(* IEC 61131-3 sources: iolistgen/src/POUs/PRG_Main, 2 files *)

(* ---- PRG_Main.decl.st ---- *)
// Назначение: точка входа приложения проверки сгенерированного кода (пример КНС-1, examples/kns): логика
//             станции в минимальном объёме — регулятор уровня LIC101 (тип Pid: вызов пишет логика станции,
//             контракт plc-process-lib 17.3) и хранение задания оператора в GVL_Persist (persist_extra),
//             затем вызов сгенерированного PRG_Devices. Ведущий насос упрощённо всегда Н1 (P101):
//             чередование, АВР и режимы станции — проект 02.
// Автор:      kr0nsch
// Версия:     0.2.0
// Документ:   docs/MANUAL_STEPS.md, раздел 9
PROGRAM PRG_Main
VAR
    xSpRestored : BOOL;   // задание оператора регулятора восстановлено из GVL_Persist после старта ПЛК
    xLeadAuto   : BOOL;   // ведущий насос в Auto, работает и следует заданию автоматики
END_VAR

(* ---- PRG_Main.impl.st ---- *)
// 1. Задание оператора регулятора уровня: после старта ПЛК — из энергонезависимой памяти
//    (GVL_Persist.rLIC101SpOper_m из persist_extra), дальше каждое изменение с HMI сохраняется туда же
IF NOT xSpRestored THEN
    GVL_Hmi.stLIC101Cmd.rSp_eu := GVL_Persist.rLIC101SpOper_m;
    xSpRestored := TRUE;
END_IF

// 2. Регулятор уровня LIC101: PV — уровнемер LT101, слежение и фактический выход — задание ведущего
//    насоса после его ограничений и рампы (с прошлого цикла). Насос не в Auto или стоит — регулятор следит
xLeadAuto := GVL_Devices.fbP101.xSpeedAutoActive;
GVL_Devices.fbLIC101(
    rPv_eu      := GVL_Devices.fbLT101.rValue_eu,
    xPvValid    := GVL_Devices.fbLT101.xValid,
    xTrack      := NOT xLeadAuto,
    rTrack_pct  := GVL_Devices.fbP101.rSpeedRef_pct,
    rOutAct_pct := GVL_Devices.fbP101.rSpeedRef_pct,
    stCmd       := GVL_Hmi.stLIC101Cmd,
    stCfg       := GVL_Persist.stLIC101Cfg,
    stRetain    := GVL_Persist.stLIC101Retain);
GVL_Devices.fbP101.rSpeedSpAuto_pct := GVL_Devices.fbLIC101.rOut_pct;
GVL_Persist.rLIC101SpOper_m := GVL_Hmi.stLIC101Cmd.rSp_eu;

// 3. Устройства перечня сигналов: вызовы и привязки сгенерированы iolistgen (src/POUs/Generated)
PRG_Devices();
